(* IEC 61131-3 sources: codesys-framework/txt/application/WeVe Utils (library)/TimeStamp/FB_TimeStampService/Commands, 5 files *)

(* ---- ForceNTPTimeSync.method.st ---- *)
METHOD ForceNTPTimeSync : E_TaskStatus
VAR
	E_TaskFeedback			: E_TaskStatus;
END_VAR

// --- BEGIN IMPLEMENTATION ---

ForceNTPTimeSync := E_TaskStatus.Busy;

CASE _wForceNTPTimeSyncState OF

	0:
		E_TaskFeedback := SetTimeBase(eTimeBase := E_TimeBase.Manual);

		IF E_TaskFeedback = E_TaskStatus.Successful THEN
			_wForceNTPTimeSyncState := _wForceNTPTimeSyncState + 10;
		ELSIF E_TaskFeedback = E_TaskStatus.Failed THEN
			_wForceNTPTimeSyncState := 100;
		END_IF

	10:
		E_TaskFeedback := SetTimeBase(eTimeBase := E_TimeBase.NTP);

		IF E_TaskFeedback = E_TaskStatus.Successful THEN
			_wForceNTPTimeSyncState := _wForceNTPTimeSyncState + 10;
		ELSIF E_TaskFeedback = E_TaskStatus.Failed THEN
			_wForceNTPTimeSyncState := 100;
		END_IF

	20:
		ForceNTPTimeSync := E_TaskStatus.Successful;
		_wForceNTPTimeSyncState := 0;

	100:
		ForceNTPTimeSync := E_TaskStatus.Failed;
		_wForceNTPTimeSyncState := 0;

END_CASE

(* ---- SetLocalTime.method.st ---- *)
METHOD SetLocalTime : E_TaskStatus
VAR_INPUT
	uiYear 					: UINT;
	uiMonth 				: UINT;
	uiDay 					: UINT;
	uiHour 					: UINT;
	uiMinute 				: UINT;
	uiSecond 				: UINT;
END_VAR
VAR
	_uliParWrite			: ULINT;
END_VAR

// --- BEGIN IMPLEMENTATION ---

_dtSetDateAndTime := DTU.DTConcat(
						uiYear := uiYear,
						uiMonth := uiMonth,
						uiDay := uiDay,
						uiHour := uiHour,
						uiMinute := uiMinute,
						uiSecond := uiSecond,
						peError := ADR(_eError)
					);

_uliParWrite:=(DT_TO_ULINT(_dtSetDateAndTime)-946684800)*1000000000;	//Compensation for 1/1/1970 vs 1/1/2000

SetLocalTime := WriteParameter(
	wIndex		:= 	16#245C,
	bySubIndex	:= 	2,
	udiTimeOut	:= 	1000,
	pDataBuffer	:=	ADR(_uliParWrite) ,
	udiDataSize	:=	8
);

(* ---- SetLocalTimeZone.method.st ---- *)
METHOD SetLocalTimeZone : E_TaskStatus
VAR_INPUT
	eTimeZone	: E_TimeZone;
END_VAR

// --- BEGIN IMPLEMENTATION ---

SetLocalTimeZone := WriteParameter(
	wIndex		:= 	16#245C,
	bySubIndex	:= 	1,
	udiTimeOut	:= 	1000,
	pDataBuffer	:=	ADR(eTimeZone) ,
	udiDataSize	:=	2
);

(* ---- SetTimeBase.method.st ---- *)
METHOD SetTimeBase :  E_TaskStatus
VAR_INPUT
	eTimeBase	: E_TimeBase;
END_VAR

// --- BEGIN IMPLEMENTATION ---

SetTimeBase := WriteParameter(
	wIndex		:= 	16#245B,
	bySubIndex	:= 	1,
	udiTimeOut	:= 	1000,
	pDataBuffer	:=	ADR(eTimeBase) ,
	udiDataSize	:=	1
);

(* ---- SetTimeServer.method.st ---- *)
METHOD SetTimeServer : E_TaskStatus
VAR_INPUT
END_VAR

// --- BEGIN IMPLEMENTATION ---
